Fanuc KAREL source: kt00580.KL

-- PROVISIONAL review KL for V1013-1; original PC SHA256 76e9b6b406d164133128fd57ff4541b5f4cf7408e0f68d5534c4afefa0d05da7
-- Incomplete behavior may be omitted. Consult companion uncertainty JSON. Do not deploy.
PROGRAM KT00580
%NOLOCKGROUP
VAR
  I2 : INTEGER
-- UNRESOLVED_DECL V1 type=000013
-- UNRESOLVED_DECL OUT type=000013
BEGIN
  -- UNRESOLVED_PC offsets 5-20; opcodes 2E,22,32,35
  -- UNRESOLVED_PC offsets 25-36; opcodes 2E,23
  -- UNRESOLVED_PC offsets 41-63; opcodes 49,21,8D,4A
  -- UNRESOLVED_PC offsets 68-72; opcodes 7F
END KT00580
